// TIA Portal V20 program export: 0 tag tables, 1 data types, 1 data blocks, 6 code blocks (in call order from the OBs), 1 instance data blocks

TYPE "zzE2eUdtA"
// stored: IsFailsafeCompliant false
   STRUCT
      m1 : Int;
      m2 : Bool;
      m3 : Int;
   END_STRUCT;
END_TYPE

DATA_BLOCK "zzE2eDb"   // DB14
{ S7_Optimized_Access := 'TRUE' }
VERSION : 0.1
// stored: AutoNumber true, DBAccessibleFromOPCUA true, DBAccessibleFromWebserver true, IsOnlyStoredInLoadMemory false, IsRetainMemResEnabled false, IsWriteProtectedInAS false, MemoryReserve 100
   VAR
      speed : Int := 150;
      dev1 { S7_SetPoint := 'True'} : "zzE2eUdtA";
   END_VAR
BEGIN
   dev1.m1 := 5;
   dev1.arr[1] := 4;
END_DATA_BLOCK

ORGANIZATION_BLOCK "Jumps"   // OB1, LAD, ProgramCycle
{ S7_Optimized_Access := 'TRUE' }
VERSION : 0.1
// stored: AutoNumber true, IsIECCheckEnabled true, SetENOAutomatically false
   VAR_INPUT
      Initial_Call : Bool;
   END_VAR
   VAR_TEMP
      valA : DInt;
      valB : DInt;
      valC : DInt;
      result : DInt;
      selector : USInt;
      caseA : USInt;
      caseB : USInt;
      done : Bool;
   END_VAR
BEGIN

REGION Network 1: Switch
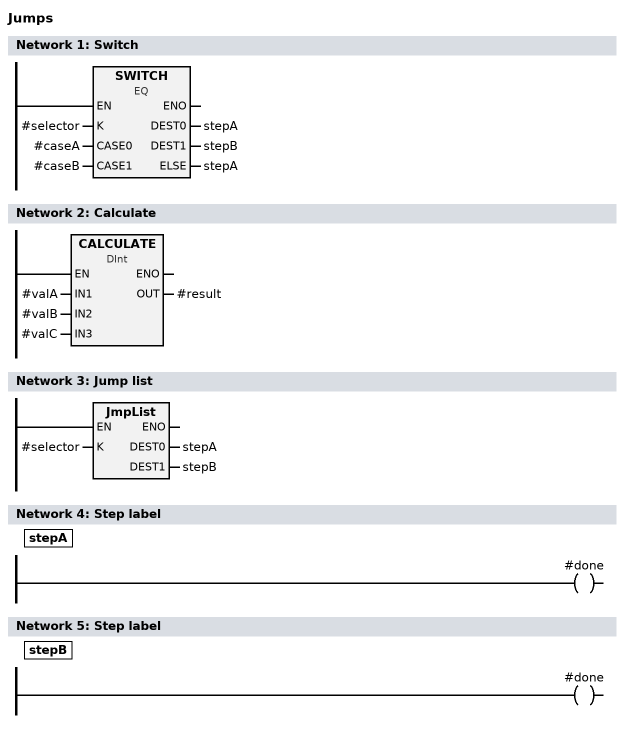
   // no SCL statement known for Switch: written as a call
   Switch(k := #selector, case0 := #caseA, case1 := #caseB, dest0 => stepA, dest1 => stepB, "else" => stepA);
END_REGION

REGION Network 2: Calculate
   RUNG wire#powerrail
      { S7_Templates := "SrcType := DInt"; S7_Expression := "(IN1 + IN2) * (IN1 - IN2)" } Calculate(in1 := #valA, in2 := #valB, in3 := #valC, out => #result)
   END_RUNG
   // the same network as SCL:
   #result := (#valA + #valB) * (#valA - #valB);
END_REGION

REGION Network 3: Jump list
   // no SCL statement known for JmpList: written as a call
   JmpList(k := #selector, dest0 => stepA, dest1 => stepB);
END_REGION

REGION Network 4: Step label
   Label( stepA )
   RUNG wire#powerrail
      Coil( #done )
   END_RUNG
   // the same network as SCL:
   stepA:
   #done := TRUE;
END_REGION

REGION Network 5: Step label
   Label( stepB )
   RUNG wire#powerrail
      Coil( #done )
   END_RUNG
   // the same network as SCL:
   stepB:
   #done := TRUE;
END_REGION
END_ORGANIZATION_BLOCK

FUNCTION_BLOCK "zzLadControl"   // FB5, LAD
{ S7_Optimized_Access := 'TRUE' }
VERSION : 0.1
// Inventory: Program control operations
// stored: AutoNumber true, IsIECCheckEnabled false, IsRetainMemResEnabled false, MemoryReserve 100, SetENOAutomatically false, UDAEnableTagReadback false
BEGIN

REGION Network 1: CoilRetValue
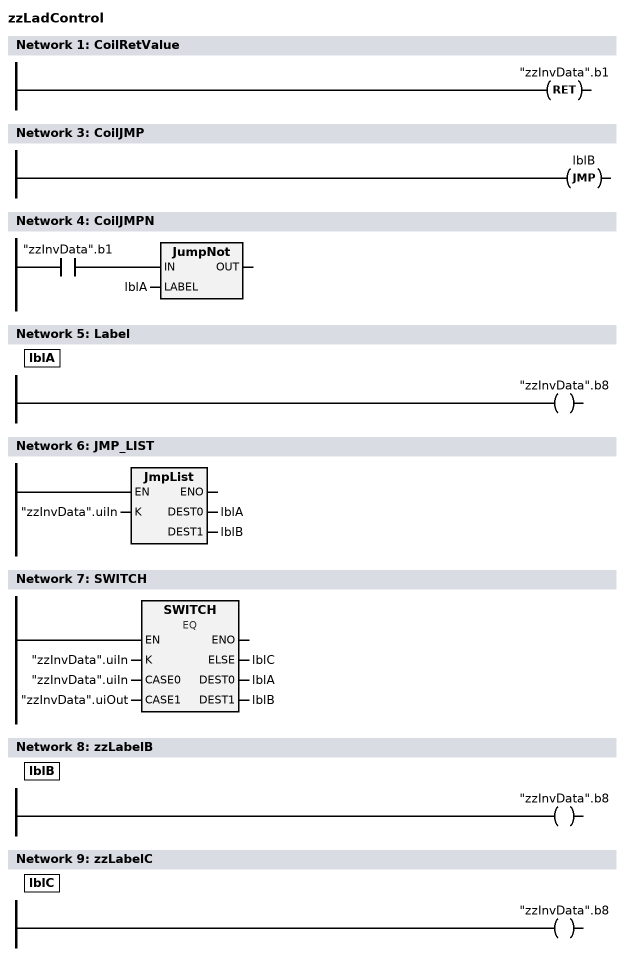
   ENO := "zzInvData".b1;
   RETURN;
END_REGION

REGION Network 2: Empty
END_REGION

REGION Network 3: CoilJMP
   RUNG wire#powerrail
      JumpCoil( lblB )
   END_RUNG
   // the same network as SCL:
   GOTO lblB;
END_REGION

REGION Network 4: CoilJMPN
   // no SCL statement known for JumpNot: written as a call
   JumpNot(in := "zzInvData".b1, label := lblA);
END_REGION

REGION Network 5: Label
   Label( lblA )
   RUNG wire#powerrail
      Coil( "zzInvData".b8 )
   END_RUNG
   // the same network as SCL:
   lblA:
   "zzInvData".b8 := TRUE;
END_REGION

REGION Network 6: JMP_LIST
   // no SCL statement known for JmpList: written as a call
   JmpList(k := "zzInvData".uiIn, dest0 => lblA, dest1 => lblB);
END_REGION

REGION Network 7: SWITCH
   // no SCL statement known for Switch: written as a call
   Switch(k := "zzInvData".uiIn,
          case0 := "zzInvData".uiIn,
          case1 := "zzInvData".uiOut,
          "else" => lblC,
          dest0 => lblA,
          dest1 => lblB);
END_REGION

REGION Network 8: zzLabelB
   Label( lblB )
   RUNG wire#powerrail
      Coil( "zzInvData".b8 )
   END_RUNG
   // the same network as SCL:
   lblB:
   "zzInvData".b8 := TRUE;
END_REGION

REGION Network 9: zzLabelC
   Label( lblC )
   RUNG wire#powerrail
      Coil( "zzInvData".b8 )
   END_RUNG
   // the same network as SCL:
   lblC:
   "zzInvData".b8 := TRUE;
END_REGION
END_FUNCTION_BLOCK

FUNCTION_BLOCK "zzBenSclColours"   // FB260, SCL
{ S7_Optimized_Access := 'TRUE' }
VERSION : 0.1
// stored: AutoNumber true, IsIECCheckEnabled false, IsRetainMemResEnabled false, MemoryReserve 100, SetENOAutomatically false, UDAEnableTagReadback false
   VAR_INPUT
      inEnable : Bool;
      inMode : Int;
      inSetpoint : Real;
   END_VAR
   VAR_OUTPUT
      outActive : Bool;
      outCount : DInt;
      outText : String[40];
   END_VAR
   VAR_IN_OUT
      ioTotal : DInt;
      ioVar : Variant;
   END_VAR
   VAR
      instColFb { S7_SetPoint := 'True'} : "zzBenSclColFb";
      instDelay { S7_SetPoint := 'True'} : TON_TIME;
      statWord : Word;
      statByte : Byte;
      statValues : Array[0..9] of Int;
      statReal : Real;
      statTime : Time;
      statDate : Date;
      statTod : Time_Of_Day;
      statChar : Char;
      statWide : WString[20];
      statFlag : Bool;
      statResult : Int;
      statTimer { S7_SetPoint := 'True'} : IEC_TIMER;
      statÄnderung : Int;
      statÜbung : Int;
   END_VAR
   VAR_TEMP
      tmpI : Int;
      tmpSum : DInt;
      tmpBit : Bool;
   END_VAR
   VAR CONSTANT
      LAST : Int := 9;
   END_VAR
BEGIN
   REGION Constants of each form
       // A line comment on a line of its own
       #statFlag := TRUE;
       #statResult := 42;
       #statResult := -8#17;
       #statWord := 16#00FF;
       #statByte := 2#1010_0101;
       #statReal := 3.14;
       #statReal := 1.5E-3;
       #statTime := T#1s_200ms;
       #statDate := D#2026-11-20;
       #statTod := TOD#12:30:00;
       #statChar := 'A';
       #outText := 'a string with // and (* inside';
       #statWide := WSTRING#'wide';
       #tmpSum := DINT#-7;
       #statWord := WORD#16#0F0F;
   END_REGION

   REGION Operands
       (* A block comment
          over two lines *)
       #outActive := #inEnable AND "zzMcTag1"; // a comment after code
       "zzBenSclColDb".motor.speed := #inMode;
       "zzBenSclColDb".values[#tmpI] := #statValues[LAST];
       #tmpBit := #statWord.%X3;
       #statByte := #statWord.%B0;
       #ioTotal += #outCount;
       "zzMcTag1" := #tmpBit;
   END_REGION

   REGION Keywords
       IF #inMode = 1 THEN
           #statResult := 1;
       ELSIF #inMode > 1 AND #inMode <= 5 THEN
           #statResult := #inMode MOD 2;
       ELSE
           #statResult := 0;
       END_IF;

       CASE #inMode OF
           0:
               #outText := 'idle';
           1..3, 5:
               #outText := 'run';
           ELSE
               #outText := '';
       END_CASE;

       #tmpSum := 0;
       FOR #tmpI := 0 TO #LAST BY 1 DO
           IF #statValues[#tmpI] < 0 THEN
               CONTINUE;
           END_IF;
           #tmpSum := #tmpSum + #statValues[#tmpI];
           IF #tmpSum > 1000 THEN
               EXIT;
           END_IF;
       END_FOR;

       #tmpI := 0;
       WHILE #tmpI < #LAST AND NOT #statFlag DO
           #tmpI := #tmpI + 1;
       END_WHILE;

       REPEAT
           #tmpI := #tmpI - 1;
       UNTIL #tmpI <= 0 OR #statFlag XOR #tmpBit
       END_REPEAT;
   END_REGION

   REGION Calls
       // An instruction with an instance and without, an FC, an FB as a multi-instance and with its DB
       #instDelay(IN := #inEnable,
                  PT := T#5s,
                  Q => #statFlag,
                  ET => #statTime);
       #statResult := MAX(IN1 := #statResult, IN2 := 10);
       #statReal := SQRT(ABS(#inSetpoint)) ** 2.0;
       #statResult := "zzBenSclColFc"(inA := #statResult, inB := 5);
       #instColFb(inStart := #statFlag,
                  outDone => #tmpBit);
       "zzBenSclColFbDb"(inStart := #inEnable);
       #outCount := INT_TO_DINT(#statResult) * 2 - #tmpSum / 3;
   END_REGION

   REGION Settled by TIA // a comment on the region's line
       (/*A multilingual comment in code*/)
       ENO := FALSE;
       IF TypeOf(#ioVar) = Int THEN
           #statÄnderung := 1;
       ELSIF TypeOf(#ioVar) = zzBenSclColType THEN
           #statÄnderung := 2;
       END_IF;
       #statTimer.TON(IN := #inEnable, PT := T#2s);
       #statÜbung := #statÄnderung + 1;
   END_REGION

   IF NOT #inEnable THEN
       GOTO lblEnd;
   END_IF;
   #outActive := #instColFb.outDone OR "zzBenSclColFbDb".outDone;
   RETURN;
   lblEnd: #outActive := FALSE;
END_FUNCTION_BLOCK

FUNCTION_BLOCK "zzE2eFbd"   // FB7, FBD
{ S7_Optimized_Access := 'TRUE' }
VERSION : 0.1
// stored: AutoNumber true, IsIECCheckEnabled false, IsRetainMemResEnabled false, MemoryReserve 100, SetENOAutomatically false, UDAEnableTagReadback false
   VAR_INPUT
      ina : Bool;
      inb : Bool;
      inc : Bool;
      ind : Bool;
      iv1 : Int;
      iv2 : Int;
   END_VAR
   VAR_OUTPUT
      outq : Bool;
      outr : Bool;
      ov1 : Int;
   END_VAR
BEGIN

REGION Network 1: And gate
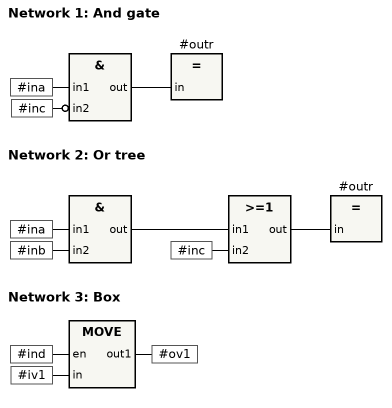
   #outr := #ina AND NOT #inc;
END_REGION

REGION Network 2: Or tree
   #outr := (#ina AND #inb) OR #inc;
END_REGION

REGION Network 3: Box
   IF #ind THEN #ov1 := #iv1; END_IF;
END_REGION
END_FUNCTION_BLOCK

FUNCTION_BLOCK "zzBenTimers"   // FB240, LAD
{ S7_Optimized_Access := 'TRUE' }
VERSION : 0.1
// Benchmark networks, timers, counters, edges
// stored: AutoNumber true, IsIECCheckEnabled false, IsRetainMemResEnabled false, MemoryReserve 100, SetENOAutomatically false, UDAEnableTagReadback false
   VAR_INPUT
      inAuto : Bool;
      inLevel : Int;
      inManual : Bool;
      inSensorA : Bool;
      inSpeed : Int;
      inStart : Bool;
   END_VAR
   VAR_OUTPUT
      outQ1 : Bool;
      outQ2 : Bool;
      outQ3 : Bool;
      outQ4 : Bool;
   END_VAR
   VAR
      instCtu { S7_SetPoint := 'True'} : CTU_INT;
      instCtuA { S7_SetPoint := 'True'} : CTU_INT;
      instTonA { S7_SetPoint := 'True'} : TON_TIME;
      instTonB { S7_SetPoint := 'True'} : TON_TIME;
      statEdge : Bool;
      statElapsed : Time;
      statHold : Bool;
      statStep : Int;
   END_VAR
   VAR_TEMP   // added for the SCL form of the ladder/FBD networks
      _w1 : Bool;
   END_VAR
BEGIN

REGION Network 1: 14 Counter with fed pins
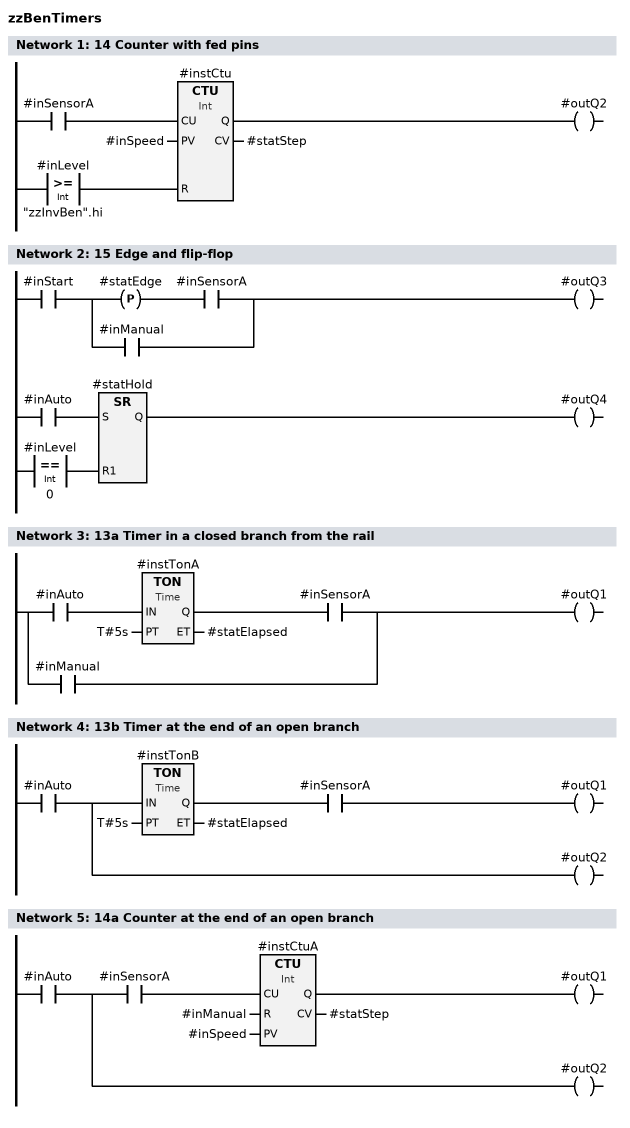
   RUNG wire#powerrail
      Contact( #inSensorA )
      { S7_Templates := "value_type := Int" } #instCtu.CTU(pv := #inSpeed, cv => #statStep, r := wire#w1)
      Coil( #outQ2 )
   END_RUNG
   RUNG wire#powerrail
      { S7_Templates := "SrcType := Int" } GE_Contact(in1 := #inLevel, in2 := "zzInvBen".hi)
   END_RUNG wire#w1
   // the same network as SCL:
   #instCtu(CU := #inSensorA, PV := #inSpeed, R := #inLevel >= "zzInvBen".hi, CV => #statStep);   // CTU
   #outQ2 := #instCtu.Q;
END_REGION

REGION Network 2: 15 Edge and flip-flop
   RUNG wire#powerrail
      Contact( #inStart )
      wire#w1
      P_Trig( #statEdge )
      Contact( #inSensorA )
      wire#w2
      Coil( #outQ3 )
   END_RUNG
   RUNG wire#w1
      Contact( #inManual )
   END_RUNG wire#w2
   RUNG wire#powerrail
      Contact( #inAuto )
      S_SR(operand := #statHold, r1 := wire#w3)
      Coil( #outQ4 )
   END_RUNG
   RUNG wire#powerrail
      { S7_Templates := "SrcType := Int" } EQ_Contact(in1 := #inLevel, in2 := 0)
   END_RUNG wire#w3
   // the same network as SCL:
   #_w1 := #inStart AND NOT #statEdge;   // rising edge
   #statEdge := #inStart;
   #outQ3 := (#_w1 AND #inSensorA) OR (#inStart AND #inManual);
   IF #inAuto THEN
       #statHold := TRUE;   // SR flip-flop
   END_IF;
   IF #inLevel = 0 THEN #statHold := FALSE; END_IF;
   #outQ4 := #statHold;
END_REGION

REGION Network 3: 13a Timer in a closed branch from the rail
   RUNG wire#powerrail
      Contact( #inAuto )
      { S7_Templates := "time_type := Time" } #instTonA.TON(pt := T#5s, et => #statElapsed)
      Contact( #inSensorA )
      wire#w1
      Coil( #outQ1 )
   END_RUNG
   RUNG wire#powerrail
      Contact( #inManual )
   END_RUNG wire#w1
   // the same network as SCL:
   #instTonA(IN := #inAuto, PT := T#5s, ET => #statElapsed);   // TON
   #outQ1 := (#instTonA.Q AND #inSensorA) OR #inManual;
END_REGION

REGION Network 4: 13b Timer at the end of an open branch
   RUNG wire#powerrail
      Contact( #inAuto )
      wire#w1
      { S7_Templates := "time_type := Time" } #instTonB.TON(pt := T#5s, et => #statElapsed)
      Contact( #inSensorA )
      Coil( #outQ1 )
   END_RUNG
   RUNG wire#w1
      Coil( #outQ2 )
   END_RUNG
   // the same network as SCL:
   #instTonB(PT := T#5s, IN := #inAuto, ET => #statElapsed);   // TON
   #outQ1 := #instTonB.Q AND #inSensorA;
   #outQ2 := #inAuto;
END_REGION

REGION Network 5: 14a Counter at the end of an open branch
   RUNG wire#powerrail
      Contact( #inAuto )
      wire#w1
      Contact( #inSensorA )
      { S7_Templates := "value_type := Int" } #instCtuA.CTU(r := #inManual, pv := #inSpeed, cv => #statStep)
      Coil( #outQ1 )
   END_RUNG
   RUNG wire#w1
      Coil( #outQ2 )
   END_RUNG
   // the same network as SCL:
   #instCtuA(CU := #inAuto AND #inSensorA, R := #inManual, PV := #inSpeed, CV => #statStep);   // CTU
   #outQ1 := #instCtuA.Q;
   #outQ2 := #inAuto;
END_REGION
END_FUNCTION_BLOCK

FUNCTION_BLOCK "zzE2eFbI"   // FB247, LAD
{ S7_Optimized_Access := 'TRUE' }
VERSION : 0.1
// stored: AutoNumber true, IsIECCheckEnabled false, IsRetainMemResEnabled false, MemoryReserve 100, SetENOAutomatically false, UDAEnableTagReadback false
   VAR_INPUT
      inV : Int;
      inW : Int;
   END_VAR
   VAR
      stV : Int := 1;
      stU { S7_SetPoint := 'True'} : "zzE2eUdtA";
   END_VAR
BEGIN

REGION Network 1
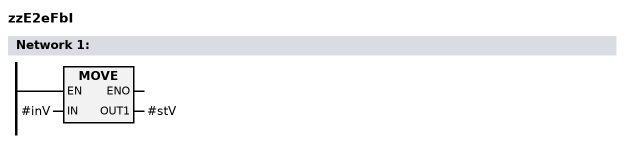
   RUNG wire#powerrail
      Move(in := #inV, out1 => #stV)
   END_RUNG
   // the same network as SCL:
   #stV := #inV;
END_REGION
END_FUNCTION_BLOCK

DATA_BLOCK "zzE2eFbI_DB"   // DB16
VERSION : 0.1
// stored: AutoNumber true, DBAccessibleFromOPCUA true, DBAccessibleFromWebserver true, InstanceOfName zzE2eFbI, InstanceOfType FB
"zzE2eFbI"
BEGIN
   stU.as[*].x := 1;   // as x
END_DATA_BLOCK
